Staubli VAL3: MoveC.pgx

public program MoveC(pointRx x_pPoint1, pointRx x_pPoint2, tool x_tTool, mdesc x_mSpeed, num& x_nMoveId)
// // 圆弧运动movec程序
// // 用该程序替代原val3程序中的movec()指令即可
// // 因为原move指令有返回值moveID，所以这里引入一个x_nMoveId，随参考传递出来
begin
  // ---------------------------------------------------------------------------- //
  // 圆弧运动movec程序
  // 用该程序替代原val3程序中的movec()指令即可
  // 因为原move指令有返回值moveID，所以这里引入一个x_nMoveId，随参考传递出来
  // ---------------------------------------------------------------------------- //
  //
  //
  x_nMoveId=movec(x_pPoint1,x_pPoint2,x_tTool,x_mSpeed)
  // log
  call logMoveMsgC(x_pPoint1,x_pPoint2,x_tTool,x_mSpeed,x_nMoveId)

end
